(* IEC 61131-3 sources: codesys-to-s7/tests/corpus/C2S7-POU-INCONST/neg, 1 file *)

(* ---- input.st ---- *)
FUNCTION_BLOCK FB_Case
VAR_INPUT
    k : INT;
END_VAR
VAR
    a : INT;
END_VAR
a := k;
END_FUNCTION_BLOCK
